(* IEC 61131-3 sources: plc-iiot-stack/src/POUs/Iiot/F_IiotTopic, 2 files *)

(* ---- F_IiotTopic.decl.st ---- *)
// Назначение: полный топик <префикс>/<хвост>; пустой префикс — только хвост. Не помещается в
//             MQTT_TOPIC_LEN — пустая строка (вызывающий считает это ошибкой).
// Автор:      kr0nsch
// Версия:     0.1.0
// Документ:   docs/plc_mqtt.md, раздел «Топики»
FUNCTION F_IiotTopic : STRING(GVL_Const.MQTT_TOPIC_LEN)
VAR_INPUT
    sPrefix : STRING(GVL_Const.IIOT_PREFIX_LEN);   // site/area/unit
    sPath : STRING(GVL_Const.MQTT_TOPIC_LEN);      // device/metric, device/alarm/suffix ...
END_VAR

(* ---- F_IiotTopic.impl.st ---- *)
IF LEN(sPrefix) = 0 THEN
    F_IiotTopic := sPath;
ELSIF LEN(sPrefix) + LEN(GVL_Const.TOPIC_SEPARATOR) + LEN(sPath) > UINT_TO_INT(GVL_Const.MQTT_TOPIC_LEN) THEN
    F_IiotTopic := '';
ELSE
    F_IiotTopic := CONCAT(CONCAT(sPrefix, GVL_Const.TOPIC_SEPARATOR), sPath);
END_IF
